Fanuc KAREL source: KB00036.KL

PROGRAM KB00036
%NOLOCKGROUP
VAR
  P1: JOINTPOS
  P2: REAL
  P3: INTEGER
BEGIN
  P2 = 1.0
  P3 = 1
  CNV_JPOS_REL(P1, P2, P3)
END KB00036
